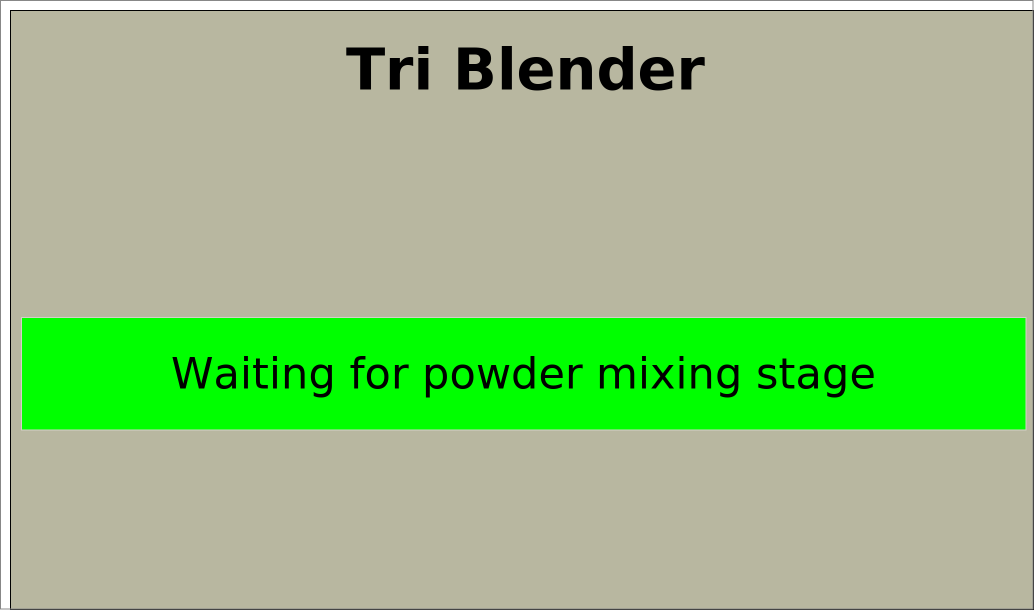
VISUALIZATION StartVisu  // 1034x610
    Rectangle (10,10 1024x600)
    Textfield (19,21 1013x96), "Tri Blender"
    Textfield (21,317 1005x113), "Waiting for powder mixing stage"
END_VISUALIZATION

// ---- 03 Project/22 InterConnection/00 General/TextList_TriBlenderUsage.TcTLO
TEXTLIST TextList_TriBlenderUsage
  0 = 'Not in Use'
  1 = 'Marinada T1'
  2 = 'Marinada T2'
  3 = 'Marinada Stanbdy'
  4 = 'Color T3'
  5 = 'Color T4'
  6 = 'Color Standby'
   = ''
END_TEXTLIST

// ---- 03 Project/22 InterConnection/00 General/vis_FB_InterConnection.TcVIS
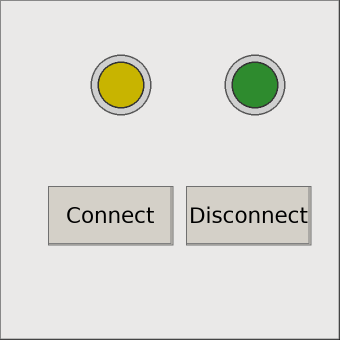
VISUALIZATION vis_FB_InterConnection  // 340x340
VAR_IN_OUT
	fb: FB_InterConnection;

END_VAR
    Rectangle (0,0 340x340)
    Button (48,186 125x59), "Connect", input disabled if: NOT fb.bAvalableToConnect
        OnMouseClick: toggle fb.reqConnect
    Button (186,186 125x59), "Disconnect", input disabled if: NOT fb.bAvalableToDisconnect
        OnMouseClick: toggle fb.reqDisconnect
    Lamp1 (220,50 70x70), variable: fb.bActive, style: Lamp-Lamp1-Green
    Lamp1 (86,50 70x70), variable: fb.bAvalableToConnect, style: Lamp-Lamp1-Yellow
END_VISUALIZATION

// ---- 03 Project/22 InterConnection/00 General/vis_InterconnectionCell.TcVIS
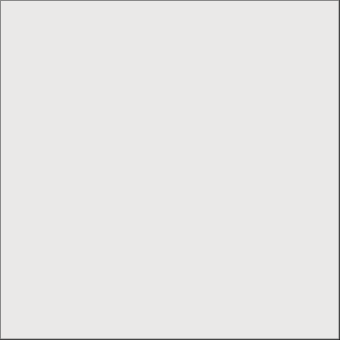
VISUALIZATION vis_InterconnectionCell  // 340x340
    Rectangle (0,0 340x340)
END_VISUALIZATION

// ---- 03 Project/22 InterConnection/00 General/vis_TriBlenderPipe.TcVIS
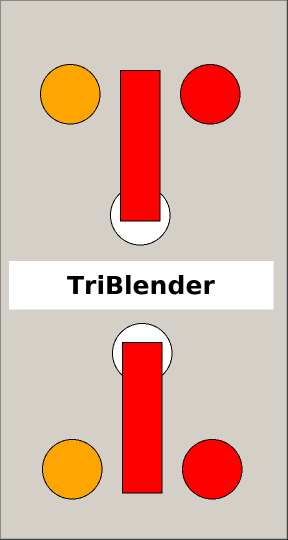
VISUALIZATION vis_TriBlenderPipe  // 288x540
    Rectangle (0,0 288x540)
    Ellipse (112,323 60x60)
        OnMouseClick: execute { eTriBlenderPipe_In:=E_TriBlenderPipe.eNone; }
    Ellipse (42,439 60x60)
        OnMouseClick: execute { eTriBlenderPipe_In:=E_TriBlenderPipe.eMarinada; }
    Ellipse (182,439 60x60)
        OnMouseClick: execute { eTriBlenderPipe_In:=E_TriBlenderPipe.eColor; }
    Ellipse (110,185 60x60)
        OnMouseClick: execute { eTriBlenderPipe_Out:=E_TriBlenderPipe.eNone; }
    Ellipse (40,64 60x60)
        OnMouseClick: execute { eTriBlenderPipe_Out:=E_TriBlenderPipe.eMarinada; }
    Ellipse (180,64 60x60)
        OnMouseClick: execute { eTriBlenderPipe_Out:=E_TriBlenderPipe.eColor; }
    RoundedRectangle (120,70 40x151), angle -30, invisible if: eTriBlenderPipe_Out<>E_TriBlenderPipe.eMarinada
        OnMouseClick: execute { eTriBlenderPipe_Out:=E_TriBlenderPipe.eNone; }
    RoundedRectangle (120,70 40x151), angle 30, invisible if: eTriBlenderPipe_Out<>E_TriBlenderPipe.eColor
        OnMouseClick: execute { eTriBlenderPipe_Out:=E_TriBlenderPipe.eNone; }
    RoundedRectangle (122,342 40x151), angle 30, invisible if: eTriBlenderPipe_In<>E_TriBlenderPipe.eMarinada
        OnMouseClick: execute { eTriBlenderPipe_In:=E_TriBlenderPipe.eNone; }
    RoundedRectangle (122,342 40x151), angle -30, invisible if: eTriBlenderPipe_In<>E_TriBlenderPipe.eColor
        OnMouseClick: execute { eTriBlenderPipe_In:=E_TriBlenderPipe.eNone; }
    Textfield (8,260 266x50), "TriBlender"
END_VISUALIZATION

// ---- 03 Project/22 InterConnection/01 Tank/TextList_E_Tank_Target.TcTLO
TEXTLIST TextList_E_Tank_Target
  0 = 'None'
  1 = 'Close'
  2 = 'Open'
  3 = 'Drain'
  4 = 'CIP'
   = ''
END_TEXTLIST

// ---- 03 Project/22 InterConnection/01 Tank/vis_FB_Tank_Target.TcVIS
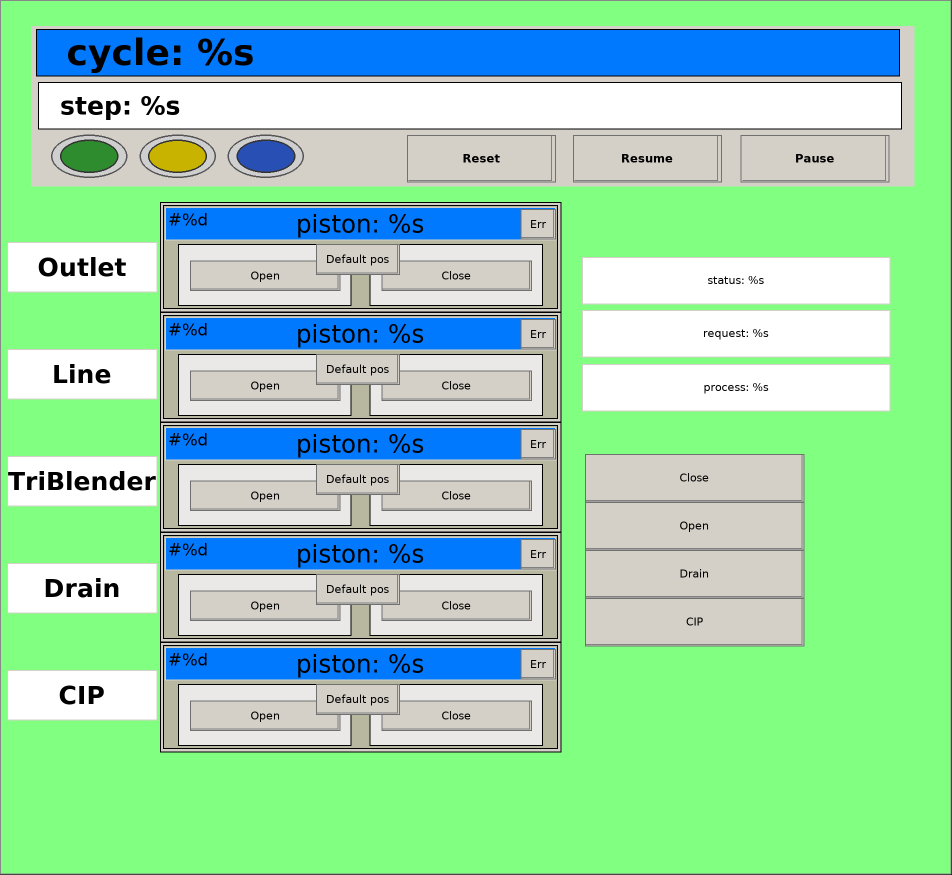
VISUALIZATION vis_FB_Tank_Target  // 952x875
VAR_IN_OUT
	fb: FB_Tank_Target;
END_VAR
    Rectangle (0,0 952x875)
    Frame (160,202 401x110)
        shows vis_Piston_Control1_Compact(stPis := fb.stPis_Outlet)
    Frame (160,312 401x110)
        shows vis_Piston_Control1_Compact(stPis := fb.stPis_Line)
    Frame (160,422 401x110)
        shows vis_Piston_Control1_Compact(stPis := fb.stPis_TriBlender)
    Frame (160,532 401x110)
        shows vis_Piston_Control1_Compact(stPis := fb.stPis_Drain)
    Frame (160,642 401x110)
        shows vis_Piston_Control1_Compact(stPis := fb.stPis_CIP)
    Frame (31,26 883x160)
        shows vis_Cycle_Control(fb := fb, sName := 'Tank Target Interface')
    Textfield (582,257 308x47), "status: %s", text variable: fb.eStatus
    Button (585,454 219x48), "Close"
        OnMouseClick: execute { fb.eReq:=E_Tank_Target.eClose; }
    Textfield (582,310 308x47), "request: %s", text variable: fb.eReq
    Textfield (582,364 308x47), "process: %s", text variable: fb.eProcess
    Button (585,502 219x48), "Open"
        OnMouseClick: execute { fb.eReq:=E_Tank_Target.eOpen; }
    Button (585,550 219x48), "Drain"
        OnMouseClick: execute { fb.eReq:=E_Tank_Target.eDrain; }
    Button (585,598 219x48), "CIP"
        OnMouseClick: execute { fb.eReq:=E_Tank_Target.eCIP; }
    Textfield (7,242 150x50), "Outlet"
    Textfield (7,349 150x50), "Line"
    Textfield (7,456 150x50), "TriBlender"
    Textfield (7,563 150x50), "Drain"
    Textfield (7,670 150x50), "CIP"
END_VISUALIZATION

// ---- 03 Project/22 InterConnection/03 Line/TextList_E_Line_Source.TcTLO
TEXTLIST TextList_E_Line_Source
  0 = 'Drain'
  1 = 'Tank_A'
  2 = 'Tank_B'
  3 = 'TapWater'
  4 = 'FillWater'
  5 = 'CIP'
   = ''
END_TEXTLIST

// ---- 03 Project/22 InterConnection/03 Line/TextList_E_Line_Target.TcTLO
TEXTLIST TextList_E_Line_Target
  0 = 'Drain'
  1 = 'Tank_A'
  2 = 'Tank_B'
  3 = 'CIP'
   = ''
END_TEXTLIST

// ---- 03 Project/23 CIP/TextList_CIP_Clients.TcTLO
TEXTLIST TextList_CIP_Clients
  0 = ' '
  1 = 'Tank1 Marinada'
  2 = 'Tank2 Marinada'
  3 = 'Tank3 Color'
  4 = 'Tank4 Color'
  5 = 'TriBlender Marinada'
  6 = 'TriBlender Color'
  7 = 'Line Marinada'
  8 = 'Line Color'
  9 = 'Local'
   = ''
END_TEXTLIST

// ---- 03 Project/23 CIP/TextList_CIP_Type.TcTLO
TEXTLIST TextList_CIP_Type
  0 = ' '
  1 = 'R Water'
  2 = 'Detergent'
  3 = 'Full'
   = ''
END_TEXTLIST

// ---- 03 Project/23 CIP/vis_CIP.TcVIS
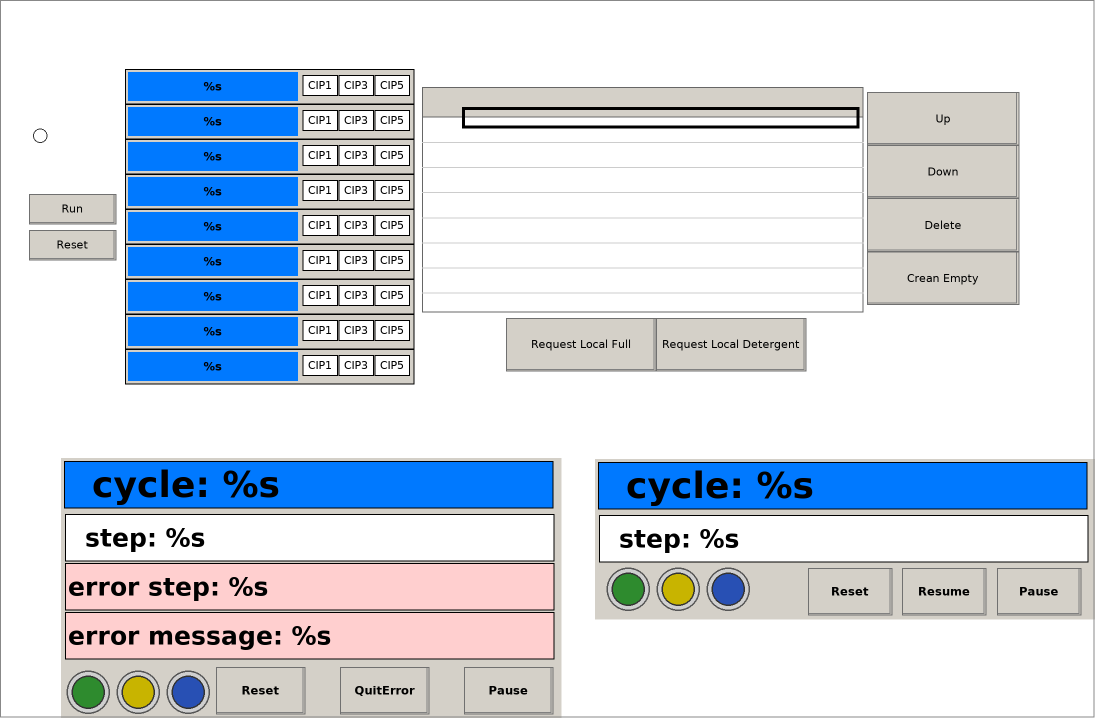
VISUALIZATION vis_CIP  // 1095x718
    Button (29,194 87x30), "Run", colour toggle: fbCIP.bRun
        toggle fbCIP.bRun
    Button (29,230 87x30), "Reset", colour toggle: fbCIP.SFCReset
        toggle fbCIP.SFCReset
    Button (506,318 150x53), "Request Local Full"
        tap fbCIP.rtReqLocalCIP_Full_HMI.CLK
    Button (656,318 150x53), "Request Local Detergent"
        tap fbCIP.rtReqLocalCIP_Detergent_HMI.CLK
    RadioButton (31,86 102x99), variable: fbCIP.eMode
        Areas[0]: Text=Off
        Areas[1]: Text=Manual
        Areas[2]: Text=Auto
    Frame (422,87 597x225)
        shows vis_CIP_ReqBuffer()
    Group (125,69 289x315)
        Frame (0,0 289x35)
            shows vis_FB_Element_CIP(fb := fbElement[E_Element_List.eTank_1])
        Frame (0,35 289x35)
            shows vis_FB_Element_CIP(fb := fbElement[E_Element_List.eTank_2])
        Frame (0,70 289x35)
            shows vis_FB_Element_CIP(fb := fbElement[E_Element_List.eTank_3])
        Frame (0,105 289x35)
            shows vis_FB_Element_CIP(fb := fbElement[E_Element_List.eTank_4])
        Frame (0,140 289x35)
            shows vis_FB_Element_CIP(fb := fbElement[E_Element_List.eTriBlender_Marinada])
        Frame (0,175 289x35)
            shows vis_FB_Element_CIP(fb := fbElement[E_Element_List.eTriBlender_Color])
        Frame (0,210 289x35)
            shows vis_FB_Element_CIP(fb := fbElement[E_Element_List.eLine_Marinada])
        Frame (0,245 289x35)
            shows vis_FB_Element_CIP(fb := fbElement[E_Element_List.eLine_Color])
        Frame (0,280 289x35)
            shows vis_FB_Element_CIP(fb := fbCIP.fbElement_Blank)
    Frame (595,459 500x160)
        shows vis_Cycle_Control(fb := fbCIP, sName := 'CIP')
    Frame (61,458 500x260)
        shows vis_Cycle_Control_1(fb := fbCIP, sName := 'CIP')
END_VISUALIZATION

// ---- 03 Project/23 CIP/vis_CIP_ReqBuffer.TcVIS
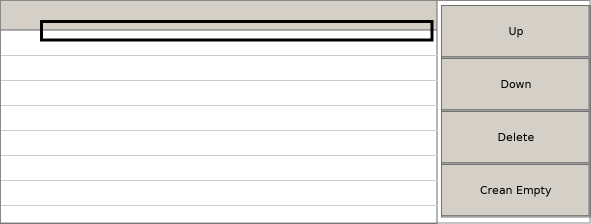
VISUALIZATION vis_CIP_ReqBuffer  // 591x224
    Table (0,0 437x224), data array: arCIP_RequestBufer
        p1137915858: fbCIP.iPosSelect_HMI
        p3854506369: arCIP_RequestBufer[INDEX].eType
        p1892666644: arCIP_RequestBufer[INDEX].eClient
    Button (441,5 150x53), "Up"
        tap fbCIP.rtPosMoveHMI_Up.CLK
    Button (441,58 150x53), "Down"
        tap fbCIP.rtPosMoveHMI_Down.CLK
    Button (441,111 150x53), "Delete"
        tap fbCIP.rtPosDeleteHMI.CLK
    Rectangle (40,20 393x21), colour toggle: fbCIP.bRun
    Button (441,164 150x53), "Crean Empty"
        tap fbCIP.rtReqCleanEmpty_HMI.CLK
END_VISUALIZATION

// ---- 03 Project/vis_Main.TcVIS
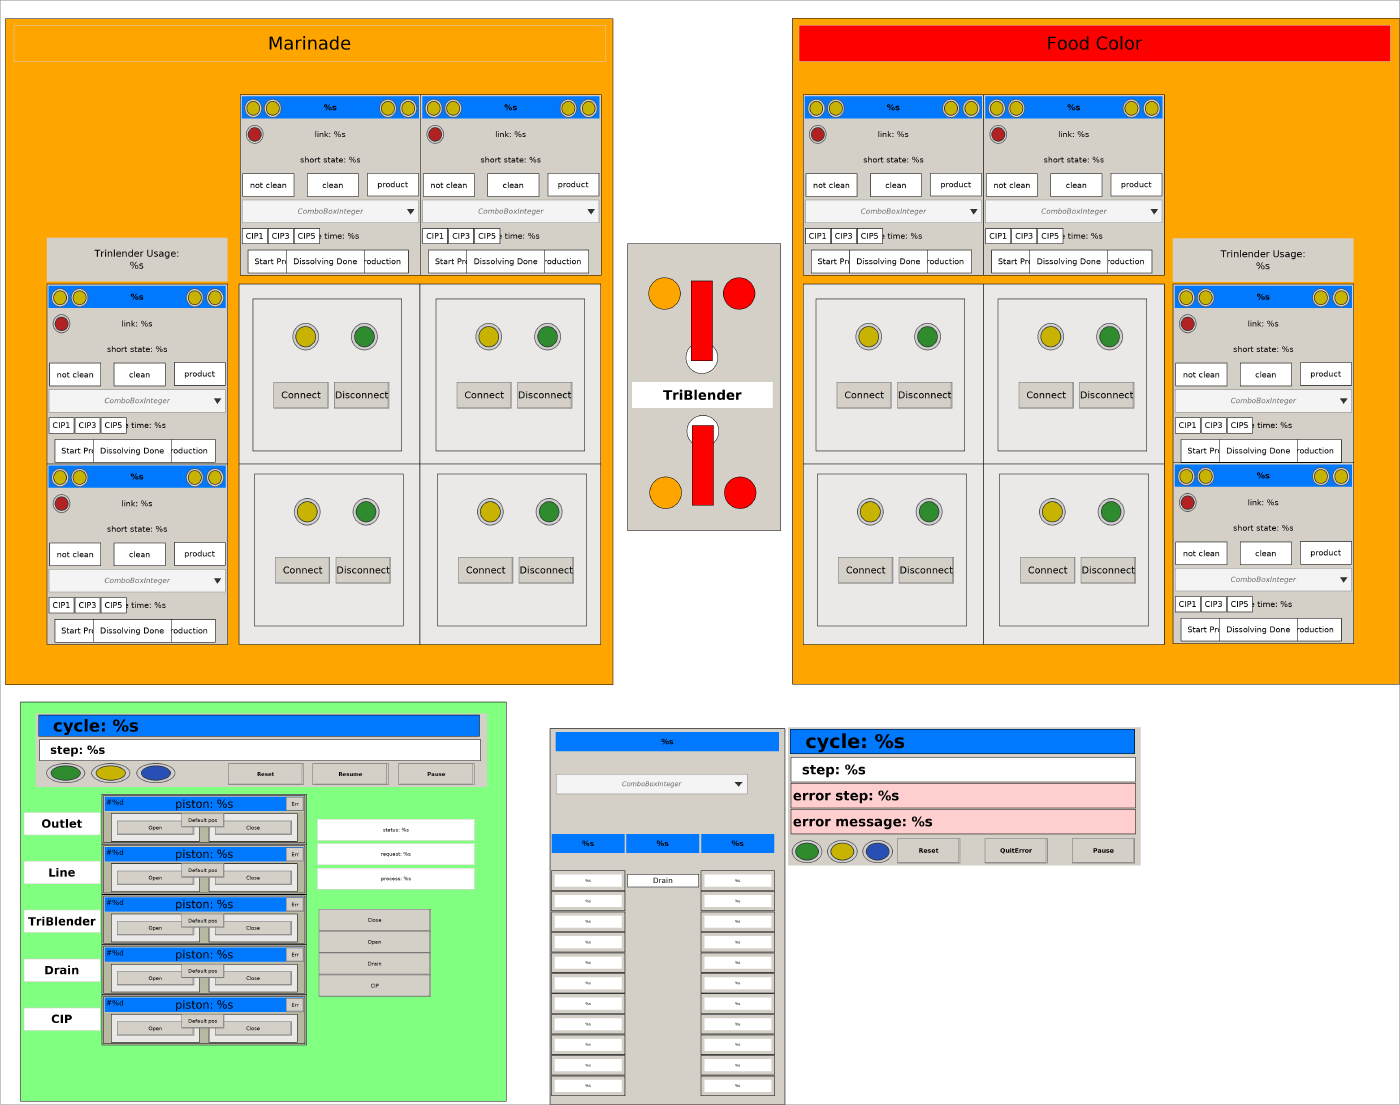
VISUALIZATION vis_Main  // 2638x2083
    Rectangle (1493,34 1145x1256)
    Frame (1513,178 341x341)
        shows vis_FB_Element(fb := fbElement[E_Element_List.eTank_3])
    Frame (1853,178 341x341)
        shows vis_FB_Element(fb := fbElement[E_Element_List.eTank_4])
    Frame (2210,535 341x341)
        shows vis_FB_Element(fb := fbElement[E_Element_List.eTriBlender_Color])
    Frame (2210,872 341x341)
        shows vis_FB_Element(fb := fbElement[E_Element_List.eLine_Color])
    Frame (1513,535 341x341)
        shows vis_InterconnectionCell()
    Frame (1853,535 341x341)
        shows vis_InterconnectionCell()
    Frame (1513,874 341x341)
        shows vis_InterconnectionCell()
    Frame (1853,874 341x341)
        shows vis_InterconnectionCell()
    Frame (1537,563 281x287)
        shows vis_FB_InterConnection(fb := fbIntCon_TriB_T3_Color)
    Frame (1880,563 281x287)
        shows vis_FB_InterConnection(fb := fbIntCon_TriB_T4_Color)
    Frame (1540,893 281x287)
        shows vis_FB_InterConnection(fb := fbIntCon_ProL_T3_Color)
    Frame (1883,893 281x287)
        shows vis_FB_InterConnection(fb := fbIntCon_ProL_T4_Color)
    Textfield (1505,47 1115x69), "Food Color"
    Group (10,35 1145x1256)
        Rectangle (0,0 1145x1256)
        Frame (442,143 341x341)
            shows vis_FB_Element(fb := fbElement[E_Element_List.eTank_1])
        Frame (782,143 341x341)
            shows vis_FB_Element(fb := fbElement[E_Element_List.eTank_2])
        Frame (78,500 341x341)
            shows vis_FB_Element(fb := fbElement[E_Element_List.eTriBlender_Marinada])
        Frame (78,839 341x341)
            shows vis_FB_Element(fb := fbElement[E_Element_List.eLine_Marinada])
        Frame (440,500 341x341)
            shows vis_InterconnectionCell()
        Frame (781,500 341x341)
            shows vis_InterconnectionCell()
        Frame (440,839 341x341)
            shows vis_InterconnectionCell()
        Frame (781,839 341x341)
            shows vis_InterconnectionCell()
        Frame (466,528 281x287)
            shows vis_FB_InterConnection(fb := fbIntCon_TriB_T1_Marin)
        Frame (811,528 281x287)
            shows vis_FB_InterConnection(fb := fbIntCon_TriB_T2_Marin)
        Frame (469,858 281x287)
            shows vis_FB_InterConnection(fb := fbIntCon_ProL_T1_Marin)
        Frame (814,858 281x287)
            shows vis_FB_InterConnection(fb := fbIntCon_ProL_T2_Marin)
        Textfield (16,12 1115x69), "Marinade"
        Textfield (78,413 340x82), "Trinlender Usage: %s", colour toggle: eTriBlenderUsage=E_TriBlenderUsage.eColor_Standby OR eTriBlenderUsage=E_TriBlenderUsage.eColor_T3 OR eTriBlenderUsage=E_TriBlenderUsage.eColor_T4, text list: 'TextList_TriBlenderUsage', text index: eTriBlenderUsage
    Textfield (2210,449 340x82), "Trinlender Usage: %s", colour toggle: eTriBlenderUsage=E_TriBlenderUsage.eMarinada_Standby OR eTriBlenderUsage=E_TriBlenderUsage.eMarinada_T1 OR eTriBlenderUsage=E_TriBlenderUsage.eMarinada_T2, text list: 'TextList_TriBlenderUsage', text index: eTriBlenderUsage
    Frame (1182,459 289x541)
        shows vis_TriBlenderPipe()
    Frame (1485,1371 664x260)
        shows vis_Cycle_Control_1(fb := fbTank1, sName := 'T1 Marinade')
    Frame (1036,1373 443x710)
        shows vis_FB_ProductionTank(fb := fbTank1)
    Frame (38,1323 916x753)
        shows vis_FB_Tank_Target(fb := fbTank1.fbTarget)
END_VISUALIZATION

// ---- GlobalTextList.TcGTLO
TEXTLIST GlobalTextList
  440 = '   message'
  1783 = '  cycle: %s'
  374 = '  step: %s'
  662 = ' %s'
  491 = '#%d'
  1694 = '%1.2f'
  153 = '%d'
  887 = '%s'
  553 = '%S'
  140 = '1/0'
  914 = '5s'
  1075 = 'Act Errors'
  1902 = 'Act State'
  690 = 'Actual'
  594 = 'Actual Errors'
  714 = 'All'
  975 = 'arCIP_RequestBufer[INDEX].eCIP_Type'
  286 = 'Auto'
  1263 = 'Axis'
  3209 = 'base time: %2.1f [sec]'
  9116 = 'ByPass'
  413 = 'bypass'
  743 = 'Cheesy Bites'
  749 = 'Cheesy Cut'
  396 = 'CIP'
  254 = 'CIP Type'
  416 = 'CIP1'
  878 = 'CIP3'
  68 = 'CIP5'
  201 = 'clean'
  677 = 'Client'
  673 = 'Close'
  1128 = 'close'
  1303 = 'Close sensor'
  8 = 'Close Sensor state'
  176 = 'Close valve'
  4398 = 'Close:'
  2046 = 'Compressor'
  520 = 'Connect'
  755 = 'Cream'
  472 = 'Crean Empty'
  742 = 'Create\nRecipe'
  1961 = 'Create Default\nRecipe'
  761 = 'Crown'
  186 = 'dealy: %.2f [sec] '
  820 = 'Default pos'
  778 = 'delay: %.2f [sec] '
  817 = 'Delete'
  713 = 'Delete\nRecipe'
  720 = 'Device 1'
  726 = 'Device 2'
  732 = 'Device 3'
  738 = 'Device 4'
  919 = 'Device Name'
  785 = 'Device State'
  178 = 'Disconnect'
  647 = 'Dissolving Done'
  47 = 'Done'
  3155 = 'Door\n#1\n'
  615 = 'Down'
  175 = 'Drain'
  460 = 'Element'
  112 = 'Emergency'
  1424 = 'Emergency Stop and Interlock'
  956 = 'EMO'
  1787 = 'Err'
  232 = 'err: %x'
  249 = 'ErrID'
  892 = 'Error'
  2981 = 'Error code: %s'
  595 = 'Error History'
  253 = 'Error Message'
  386 = 'error message: %s'
  896 = 'Error message: %s'
  5 = 'error reason: %s'
  304 = 'error step: %s'
  114 = 'Errors'
  5489 = 'Errors Search\nBuffer'
  105 = 'Errors: %d'
  3404 = 'ES Bypass'
  767 = 'Flour'
  752 = 'Food Color'
  2114 = 'Get\nLast Err'
  694 = 'History'
  756 = 'History Errors'
  3107 = 'Initialization'
  410 = 'Interlock'
  1912 = 'Interlock\nZone#1'
  4542 = 'Intilize'
  2697 = 'Last Return:'
  251 = 'Level'
  985 = 'Line'
  315 = 'link: %s'
  971 = 'Load\nRecipe'
  1122 = 'Load Recipe\nfrom file'
  135 = 'Local'
  70 = 'Main'
  2930 = 'Man'
  245 = 'Manual'
  534 = 'Marinade'
  104 = 'max: %.2f [sec] '
  11600 = 'Memo PB State'
  1148 = 'Message:'
  918 = 'min: %.2f [sec] '
  252 = 'Module Description'
  773 = 'Mozza'
  4048 = 'Mute'
  2718 = 'N'
  2076 = 'New Recipe Name:'
  920 = 'No'
  721 = 'not clean'
  181 = 'Off'
  2479 = 'OFF'
  922 = 'on'
  1164 = 'On duty: %0.1f [%]'
  952 = 'Open'
  255 = 'open'
  4392 = 'Open :'
  1663 = 'Open sensor'
  128 = 'Open Sensor state'
  197 = 'Open valve'
  779 = 'Open1'
  784 = 'Open2'
  790 = 'Open3'
  796 = 'Open4'
  444 = 'Outlet'
  1703 = 'P'
  664 = 'Password: %s'
  9135 = 'Path:'
  313 = 'Pause'
  659 = 'Pause History'
  821 = 'Piston Param'
  692 = 'piston: %s'
  704 = 'Play'
  106 = 'PLC Ver: %s'
  1953 = 'POU name: %s'
  157 = 'process: %s'
  687 = 'product'
  240 = 'Production'
  48 = 'QuitError'
  117 = 'R'
  231 = 'Ready'
  942 = 'Recipe'
  908 = 'recipe: %s'
  3336 = 'ReInit'
  2325 = 'Release ES'
  2568 = 'Reload'
  746 = 'Request Local'
  190 = 'Request Local Detergent'
  391 = 'Request Local Full'
  795 = 'request: %s'
  650 = 'Reset'
  264 = 'Reset\nErr'
  928 = 'Reset Errors'
  429 = 'Resume'
  4367 = 'Root Folder:'
  593 = 'Run'
  522 = 'Save Recipe\nto File'
  1817 = 'Save Recipe\nto file'
  1340 = 'Search'
  2084 = 'Selected Recipe:'
  2934 = 'Semi'
  1537 = 'sensor'
  183 = 'Sensor \nexist'
  814 = 'Sesame'
  953 = 'short state: %s'
  2834 = 'Standby'
  36 = 'Start Production'
  134 = 'state time: %s'
  2993 = 'state: %s'
  976 = 'status: %s'
  14674 = 'Stop\nReset All'
  812 = 'Stop Production'
  643 = 'T.C  logo '
  5392 = 'Table Index:'
  750 = 'Test'
  526 = 'Time'
  80 = 'Timing'
  1281 = 'ToBe Done'
  563 = 'TriBlender'
  96 = 'TriBlenDer'
  451 = 'Trinlender Usage:\n%s'
  915 = 'Type'
  316 = 'Up'
  745 = 'User: %s'
  810 = 'Valve'
  927 = 'Variable Name'
  936 = 'Variable Value'
  802 = 'Wet'
  808 = 'Wrap'
END_TEXTLIST
